// TIA Portal V19 export
VAR_GLOBAL   // PLC tag table "CP"
   DI_CP_Start AT %I0.4 : Bool;
   DI_CP_Stop AT %I0.5 : Bool;
   DI_CP_Reset AT %I0.6 : Bool;
   DI_CP_Auto AT %I0.7 : Bool;
   DI_CP_Manual AT %I1.0 : Bool;
   DI_CP_Request AT %I1.1 : Bool;
   DQ_CP_Start AT %Q0.0 : Bool;
   DQ_CP_Stop AT %Q0.1 : Bool;
   DQ_CP_Reset AT %Q0.2 : Bool;
   DQ_CP_Request AT %Q0.3 : Bool;
END_VAR
